            Script: ugo_update_outputs()
      Case (caseValue=14)
        Folder Unsuspending [hidden by the author, left out]
      Case (caseValue=15)
        Folder Aborting [hidden by the author, left out]
      Case (caseValue=16)
        Folder Aborted [hidden by the author, left out]
      Case (caseValue=17)
        Folder Clearing [hidden by the author, left out]
    Script: log_state(STATE_Info)
    Script: log_warning(WARNING.MSG)
    Script: log_error(ERROR.MSG)
    Folder Times [hidden by the author, left out]
    SuppressedNode
      Script: sync()
    Wait Sleep waitTime=0.1
Thread Thread_1 (runOnlyOnce=false)
  If Start_thread≟ True
    Weight_value := get_weight()
    Wait Sleep waitTime=0.1
    Script: sync()
  SuppressedNode
    If switch_spat_M≟ True (checkContinuously=true)
      If level≥10.00
        MoveJ speed 60 deg/s, acceleration 80 deg/s^2 (useActiveTCP=true) feature=Base
          Waypoint pick_spat_L_abv: TCP in base x=247.376 y=-151.301 z=298.406 mm, rx=0 ry=-0.0005 rz=3.0677 rad; joints [-4.058, -56.828, -117.366, -95.794, 90.156, 90.183] deg; TCP offset x=0 y=0 z=161 mm, rx=3.1415 ry=0 rz=0 rad
        MoveL speed 250 mm/s, acceleration 1200 mm/s^2 (useActiveTCP=true) feature=Base
          Waypoint spat_L_pick: TCP in base x=244.425 y=-151.048 z=192.288 mm, rx=0 ry=-0.0005 rz=3.0677 rad; joints [-4.109, -56.947, -132.87, -80.171, 90.162, 90.196] deg
          URCap Gripper (Robotiq_Grippers, Robotiq Inc.) dataModel(position=100.0, force=30.0, speed=0.0, positionInDouble=100.0, forceInDouble=30.0, speedInDouble=0.0, slaveIds=[9], blocking=true)
          Waypoint spat_L_lift: TCP in base x=247.5 y=-151.291 z=242.147 mm, rx=0 ry=-0.0005 rz=3.0677 rad; joints [-4.086, -56.571, -125.696, -87.721, 90.161, 90.187] deg
          Waypoint spat_L_up: TCP in base x=248.632 y=-94.371 z=425.351 mm, rx=0 ry=-0.0005 rz=3.0677 rad; joints [9.417, -57.776, -97.699, -114.51, 90.125, 103.584] deg
  SuppressedNode
    work_done := True
  SuppressedNode
    Script: sync()
SubProgram  [hidden by the author, left out]
SubProgram  [hidden by the author, left out]
SubProgram Sub_Action_V4 [hidden by the author, left out]
